FUNCTION_BLOCK VltFixtureMembers
VAR_INPUT
	bGo : BOOL;
END_VAR
VAR
	nTick : INT;
END_VAR

nTick := nTick + 1;

METHOD CfcStep : BOOL
VAR_INPUT
	bIn : BOOL;
END_VAR
END_METHOD

ACTION SfcRun:
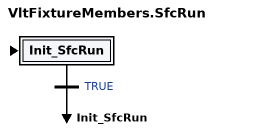
INITIAL_STEP Init_SfcRun:
END_STEP
TRANSITION FROM Init_SfcRun TO Init_SfcRun
    := TRUE;
END_TRANSITION
END_ACTION

METHOD Visible : BOOL
VAR_INPUT
	bIn : BOOL;
END_VAR
Visible := bIn;
END_METHOD

END_FUNCTION_BLOCK

(* stored: Version 1.1.0.1, ProductVersion 3.1.4024.16
   POU VltFixtureMembers: Id {631b6bc2-a4fd-47dd-9a95-80130daf31c6}, SpecialFunc None
   Method CfcStep: Id {60457d1d-8255-47dc-a7a8-a5397dc10088}
   Action SfcRun: Id {2c75a91a-3078-421b-9ba0-7bd0522653bd}
   Method Visible: Id {c8e8fa50-2b6d-4ee6-8191-46dd5571c290} *)
